Fanuc KAREL source: KO00051.KL

PROGRAM KO00051
%NOLOCKGROUP
%ENVIRONMENT MIR
VAR
  P1: XYZWPR
  P2: POSITION
  F: BOOLEAN
  OUT: XYZWPREXT
BEGIN
  F = TRUE
  OUT = MIRROR(P1, P2, F)
END KO00051
